// TIA Portal V20 export
TYPE "WT2_Vb_Status_UDT"
   STRUCT
      iHandshake : Int;
      Fehler : Struct
         bE0000_KonfigFehler : Bool;
         bE0001_Reserviert : Bool;
         bE0002_InvUngueltig : Bool;
         bE0003_Reserviert : Bool;
         bE0004_Reserviert : Bool;
         bE0005_Reserviert : Bool;
         bE0006_Reserviert : Bool;
         bE0007_KonfigFehlerKdKonst : Bool;
         bE0008_KonfigFehlerVrKonst : Bool;
         bE0009_Reserviert : Bool;
         bE0010_Reserviert : Bool;
         bE0011_Reserviert : Bool;
         bE0012_Reserviert : Bool;
         b035_Reserve : Bool;
         b036_Reserve : Bool;
         b037_Reserve : Bool;
         by04_Reserve : Byte;
         by05_Reserve : Byte;
      END_STRUCT;
      Alarm : Struct
         bA1000_Reserviert : Bool;
         bA1001_SlaveAusg : Bool;
         bA1002_Reserviert : Bool;
         bA1003_HauptMasterAusg : Bool;
         bA1004_ZuwenigVDLeistungVerf : Bool;
         bA1005_HDVerbundAusg : Bool;
         bA1006_NDVerbundAusg : Bool;
         bA1007_Reserviert : Bool;
         bA1008_Reserviert : Bool;
         bA1009_MVbMasterAktiv : Bool;
         bA1010_ObjektIDMehrfVorhanden : Bool;
         b1011_KonfigAlarmAnfVd : Bool;
         b1012_KonfigAlarmFreigabeVd : Bool;
         b075_Reserve : Bool;
         b076_Reserve : Bool;
         b077_Reserve : Bool;
         by08_Reserve : Byte;
         by09_Reserve : Byte;
      END_STRUCT;
      Zustand : Struct
         bFehlerzustandAktiv : Bool;
         bAlarmzustandAktiv : Bool;
         bSystemMeldungAktiv : Bool;
         bSeviceMeldungAktiv : Bool;
         bStopManuell : Bool;
         bStopAuto : Bool;
         bStopExtern : Bool;
         bBetriebAuto : Bool;
         bBetriebManuell : Bool;
         bAnlaufAuto : Bool;
         bAnlaufManuell : Bool;
         bManuellStoppen : Bool;
         b114_Reserve : Bool;
         b115_Reserve : Bool;
         b116_Reserve : Bool;
         b117_Reserve : Bool;
         by12_Reserve : Byte;
         bInventarAufnahme : Bool;
         bStartbefehlManuell : Bool;
         bStandbyMasterInit : Bool;
         bStandbyMasterPassiv : Bool;
         bStandbyMasterAktiv : Bool;
         bInitialisierung : Bool;
         bFreigabeWeitVdNötig : Bool;
         bAnforderungVdAktiv : Bool;
         bZuschSperreTodband : Bool;
         bBeschrLaufendeVd : Bool;
         bZuschSperreSinkenderBed : Bool;
         bLastsperreAktiv : Bool;
         bMasterGesperrt : Bool;
         bSollwertAnhebung : Bool;
         bSollwertAbsenkung : Bool;
         bPSaugTiefSperre : Bool;
         bAnfHDVerbund : Bool;
         bBoosterFreigabeFehlt : Bool;
         bAnforderungBooster : Bool;
         bHDVerbundFreigabeFehlt : Bool;
         bHDVerbundFreigabeMan : Bool;
         bBoosterFreigabeMan : Bool;
         bLeistBeschrAktiv : Bool;
         bZuschSperreLeistBesch : Bool;
         bZuschaltverzögerung : Bool;
         b161_Reserve : Bool;
         b162_Reserve : Bool;
         b163_Reserve : Bool;
         b164_Reserve : Bool;
         b165_Reserve : Bool;
         b166_Reserve : Bool;
         b167_Reserve : Bool;
         by17_Reserve : Byte;
      END_STRUCT;
      DigIn : Struct
         bStartbefehlVerbund : Bool;
         bSollwertB : Bool;
         bVerbundleistExtPlus : Bool;
         bVerbundleistExtMinus : Bool;
         bElLeistungZuHoch : Bool;
         bSollwertBHeizen : Bool;
         bUmschaltungWirksinn : Bool;
         b187_Reserve : Bool;
         by19_Reserve : Byte;
         by20_Reserve : Byte;
         by21_Reserve : Byte;
      END_STRUCT;
      DigOut : Struct
         bVerbundBereit : Bool;
         b221_Reserve : Bool;
         bFreigabeBoosterVerbund : Bool;
         bAlarmVerfLeistung : Bool;
         b224_Reserve : Bool;
         b225_Reserve : Bool;
         b226_Reserve : Bool;
         b227_Reserve : Bool;
         by23_Reserve : Byte;
         by24_Reserve : Byte;
         by25_Reserve : Byte;
      END_STRUCT;
      iAnzVd : Int;
      chRemoteSensEinheit : Char;
      chLeistRegEinheit : Char;
      rLeistRegIst : Real;
      rLeistRegSoll : Real;
      rVerbLeistSoll : Real;
      rVerbLeistSollVol : Real;
      rVerbLeistIst : Real;
      rVerbLeistIstVol : Real;
      rVeV : Real;
      rVevVol : Real;
      rVeD : Real;
      rVedVol : Real;
      rFVolMaxVerbund : Real;
      iNaechsterVdein : Int;
      iNaechsterVdaus : Int;
      rRemoteSensIst : Real;
      rVrTempEin : Real;
      rVrTempAus : Real;
      rKdrTempEin : Real;
      rKdrTempAus : Real;
      rReserveReal : Array[0..6] of Real;
      byReserveByte : Array[0..1] of Byte;
   END_STRUCT;
END_TYPE
